FUNCTION_BLOCK Stop1Coord (* Basic Function Block Type *)
  (* Standard: 61499-2 *)
  (* Version 0.0, 11/25/2026, Schneider Electric, Conveyor Stop 1 coordinator with primary Testing done and secondary sensor check *)
  PACKAGE Main;
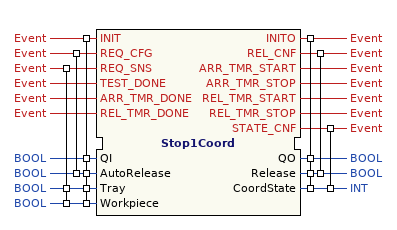
  EVENT_INPUT
    INIT WITH QI, AutoRelease, Tray, Workpiece; (* Initialization Request *)
    REQ_CFG WITH AutoRelease; (* Auto-release configuration update from Station 1 *)
    REQ_SNS WITH Tray, Workpiece; (* Stop 1 tray and workpiece sensor update *)
    TEST_DONE; (* Primary Testing pass-complete notification from Station 1 *)
    ARR_TMR_DONE; (* Tray arrival settle timer elapsed *)
    REL_TMR_DONE; (* Tray departure stopper clear delay elapsed *)
  END_EVENT
  EVENT_OUTPUT
    INITO WITH QO, Release, CoordState; (* Initialization Confirm *)
    REL_CNF WITH Release; (* Stop 1 release command update *)
    ARR_TMR_START; (* Start tray arrival settle debounce timer *)
    ARR_TMR_STOP; (* Cancel tray arrival settle debounce timer *)
    REL_TMR_START; (* Start post-departure release clear timer *)
    REL_TMR_STOP; (* Cancel post-departure release clear timer *)
    STATE_CNF WITH CoordState; (* Coordinator state update *)
  END_EVENT
  VAR_INPUT
    QI : BOOL := TRUE; (* Input event qualifier *)
    AutoRelease : BOOL := FALSE; (* Stop 1 automatic release enable from Station 1 *)
    Tray : BOOL := FALSE; (* Tray present at Stop 1 (M1.DI02) *)
    Workpiece : BOOL := FALSE; (* Workpiece present in Station 1 pocket (M1.DI05) *)
  END_VAR
  VAR_OUTPUT
    QO : BOOL; (* Output event qualifier *)
    Release : BOOL := FALSE; (* Temporary release command to Stop1 StopPoint *)
    CoordState : INT := 0; (* 0=Idle,1=ArriveSettle,2=WaitTestDone,3=WaitPartCheck,4=Releasing,5=RelClearWait *)
  END_VAR
  VAR
    state : INT := 0; (* Internal state machine value *)
    wantRelCnf : BOOL := FALSE; (* Pending REL_CNF event flag *)
    wantArrStart : BOOL := FALSE; (* Pending ARR_TMR_START event flag *)
    wantArrStop : BOOL := FALSE; (* Pending ARR_TMR_STOP event flag *)
    wantRelStart : BOOL := FALSE; (* Pending REL_TMR_START event flag *)
    wantRelStop : BOOL := FALSE; (* Pending REL_TMR_STOP event flag *)
  END_VAR
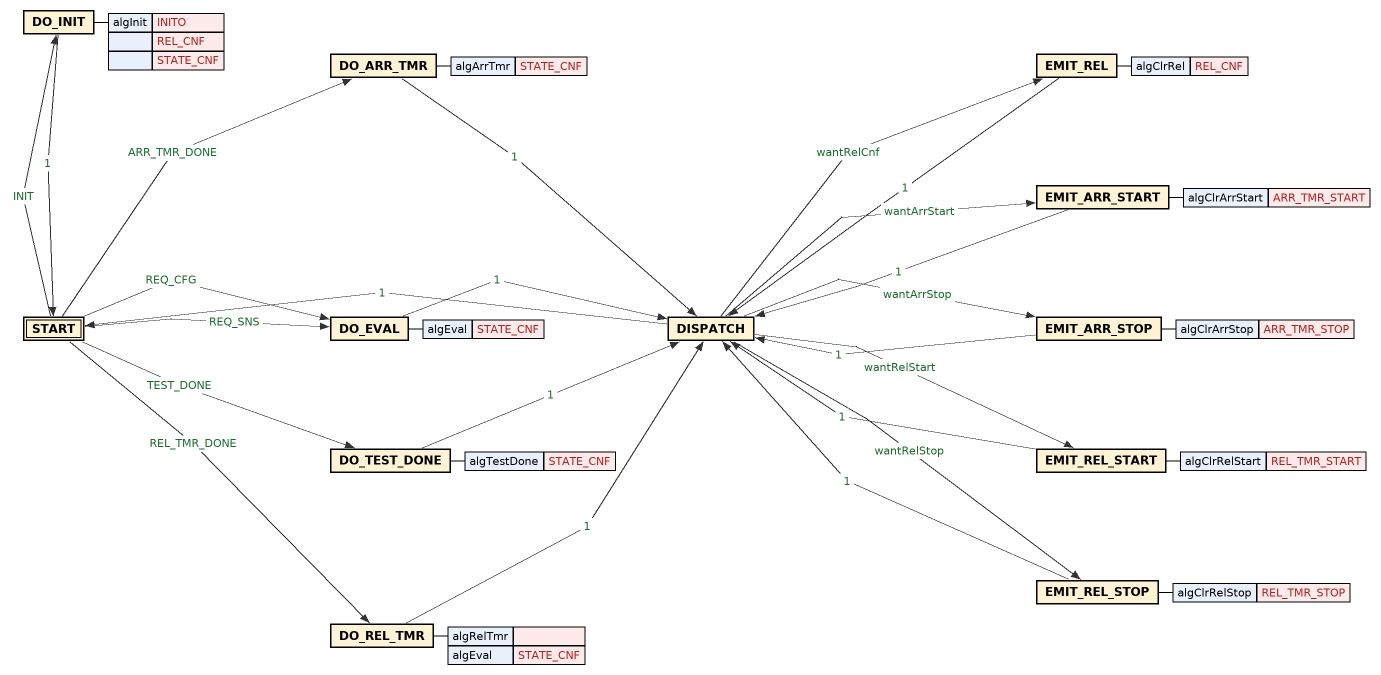
  EC_STATES
    START; (* Initial State *)
    DO_INIT : algInit -> INITO, -> REL_CNF, -> STATE_CNF;
    DO_EVAL : algEval -> STATE_CNF;
    DO_ARR_TMR : algArrTmr -> STATE_CNF;
    DO_TEST_DONE : algTestDone -> STATE_CNF;
    DO_REL_TMR : algRelTmr, algEval -> STATE_CNF;
    DISPATCH;
    EMIT_REL : algClrRel -> REL_CNF;
    EMIT_ARR_START : algClrArrStart -> ARR_TMR_START;
    EMIT_ARR_STOP : algClrArrStop -> ARR_TMR_STOP;
    EMIT_REL_START : algClrRelStart -> REL_TMR_START;
    EMIT_REL_STOP : algClrRelStop -> REL_TMR_STOP;
  END_STATES
  EC_TRANSITIONS
    START TO DO_INIT := INIT;
    DO_INIT TO START := 1;
    START TO DO_EVAL := REQ_CFG;
    START TO DO_EVAL := REQ_SNS;
    START TO DO_ARR_TMR := ARR_TMR_DONE;
    START TO DO_TEST_DONE := TEST_DONE;
    START TO DO_REL_TMR := REL_TMR_DONE;
    DO_EVAL TO DISPATCH := 1;
    DO_ARR_TMR TO DISPATCH := 1;
    DO_TEST_DONE TO DISPATCH := 1;
    DO_REL_TMR TO DISPATCH := 1;
    DISPATCH TO EMIT_REL := wantRelCnf;
    EMIT_REL TO DISPATCH := 1;
    DISPATCH TO EMIT_ARR_START := wantArrStart;
    EMIT_ARR_START TO DISPATCH := 1;
    DISPATCH TO EMIT_ARR_STOP := wantArrStop;
    EMIT_ARR_STOP TO DISPATCH := 1;
    DISPATCH TO EMIT_REL_START := wantRelStart;
    EMIT_REL_START TO DISPATCH := 1;
    DISPATCH TO EMIT_REL_STOP := wantRelStop;
    EMIT_REL_STOP TO DISPATCH := 1;
    DISPATCH TO START := 1;
  END_TRANSITIONS
  ALGORITHM algInit IN ST: (* Initialize Stop 1 coordinator state and outputs *)
QO := QI;
state := 0;
Release := FALSE;
CoordState := 0;
wantRelCnf := FALSE;
wantArrStart := FALSE;
wantArrStop := FALSE;
wantRelStart := FALSE;
wantRelStop := FALSE;
  END_ALGORITHM
  ALGORITHM algArrTmr IN ST: (* Evaluate arriving tray after arrival settle delay *)
IF AutoRelease AND (state = 1) THEN
	IF NOT Tray THEN
		state := 0;
	ELSIF Workpiece THEN
		(* Tray arrived already carrying a workpiece in pocket 1 -> bypass *)
		IF NOT Release THEN
			Release := TRUE;
			wantRelCnf := TRUE;
		END_IF;
		state := 4;
	ELSE
		(* Tray arrived empty -> wait for primary TEST_DONE from Testing *)
		state := 2;
	END_IF;
END_IF;
CoordState := state;
  END_ALGORITHM
  ALGORITHM algTestDone IN ST: (* Handle primary Testing pass-complete notification *)
IF AutoRelease THEN
	IF state = 1 THEN
		wantArrStop := TRUE;
	END_IF;
	IF (state = 1) OR (state = 2) THEN
		IF NOT Tray THEN
			state := 0;
		ELSIF Workpiece THEN
			(* Primary TEST_DONE + Secondary Tray & Workpiece confirmed *)
			IF NOT Release THEN
				Release := TRUE;
				wantRelCnf := TRUE;
			END_IF;
			state := 4;
		ELSE
			(* Primary TEST_DONE received; wait for part to land on M1.DI05 *)
			state := 3;
		END_IF;
	END_IF;
END_IF;
CoordState := state;
  END_ALGORITHM
  ALGORITHM algRelTmr IN ST: (* Clear Release after tray clears Stopper 1 *)
IF state = 5 THEN
	IF Release THEN
		Release := FALSE;
		wantRelCnf := TRUE;
	END_IF;
	state := 0;
END_IF;
  END_ALGORITHM
  ALGORITHM algEval IN ST: (* Evaluate Stop 1 release state on config or sensor changes *)
IF NOT AutoRelease THEN
	IF state = 1 THEN
		wantArrStop := TRUE;
	END_IF;
	IF state = 5 THEN
		wantRelStop := TRUE;
	END_IF;
	IF Release THEN
		Release := FALSE;
		wantRelCnf := TRUE;
	END_IF;
	state := 0;
ELSE
	IF NOT Tray THEN
		IF state = 1 THEN
			wantArrStop := TRUE;
			state := 0;
		ELSIF (state = 2) OR (state = 3) THEN
			state := 0;
		ELSIF state = 4 THEN
			wantRelStart := TRUE;
			state := 5;
		END_IF;
	ELSE
		IF state = 3 THEN
			(* Primary TEST_DONE already received -> secondary check *)
			IF Workpiece THEN
				IF NOT Release THEN
					Release := TRUE;
					wantRelCnf := TRUE;
				END_IF;
				state := 4;
			END_IF;
		ELSIF state = 0 THEN
			wantArrStart := TRUE;
			state := 1;
		END_IF;
		(* Note: in state = 2 (WaitTestDone), Workpiece alone NEVER opens the stopper! *)
	END_IF;
END_IF;

CoordState := state;
  END_ALGORITHM
  ALGORITHM algClrRel IN ST: (* Clear REL_CNF emit flag *)
wantRelCnf := FALSE;
  END_ALGORITHM
  ALGORITHM algClrArrStart IN ST: (* Clear ARR_TMR_START emit flag *)
wantArrStart := FALSE;
  END_ALGORITHM
  ALGORITHM algClrArrStop IN ST: (* Clear ARR_TMR_STOP emit flag *)
wantArrStop := FALSE;
  END_ALGORITHM
  ALGORITHM algClrRelStart IN ST: (* Clear REL_TMR_START emit flag *)
wantRelStart := FALSE;
  END_ALGORITHM
  ALGORITHM algClrRelStop IN ST: (* Clear REL_TMR_STOP emit flag *)
wantRelStop := FALSE;
  END_ALGORITHM
END_FUNCTION_BLOCK
